{attribute 'qualified_only'}
VAR_GLOBAL CONSTANT
	//This GVL contains a list of TwinCAT Errors and their corresponding error codes.
	MAX_INDEX		: INT := 744;
	
	{warning disable C0198} //disable string length warning, strings will automatically be truncated
	List			: ARRAY[0..MAX_INDEX] OF ST_TcError :=
	[
		//0 -----------------------------------
		(code		:= 0
		,message 	:= '0.  No Error')
		//1 -----------------------------------
		,(code		:= 1
		,message 	:= '1.  Internal error')
		//2 -----------------------------------
		,(code		:= 2
		,message 	:= '2.  No Rtime')
		//3 -----------------------------------
		,(code		:= 3
		,message 	:= '3.  Allocation locked memory error')
		//4 -----------------------------------
		,(code		:= 4
		,message 	:= '4.  Insert mailbox error')
		//5 -----------------------------------
		,(code		:= 5
		,message 	:= '5.  Wrong receive HMSG')
		//6 -----------------------------------
		,(code		:= 6
		,message 	:= '6.  target port not found')
		//7 -----------------------------------
		,(code		:= 7
		,message 	:= '7.  target machine not found')
		//8 -----------------------------------
		,(code		:= 8
		,message 	:= '8.  Unknown command ID')
		//9 -----------------------------------
		,(code		:= 9
		,message 	:= '9.  Bad task ID')
		//10 -----------------------------------
		,(code		:= 10
		,message 	:= '10.  No IO')
		//11 -----------------------------------
		,(code		:= 11
		,message 	:= '11.  Unknown ADS command')
		//12 -----------------------------------
		,(code		:= 12
		,message 	:= '12.  Win 32 error')
		//13 -----------------------------------
		,(code		:= 13
		,message 	:= '13.  Port not connected')
		//14 -----------------------------------
		,(code		:= 14
		,message 	:= '14.  Invalid ADS length')
		//15 -----------------------------------
		,(code		:= 15
		,message 	:= '15.  Invalid ADS Net ID')
		//16 -----------------------------------
		,(code		:= 16
		,message 	:= '16.  Low Installation level')
		//17 -----------------------------------
		,(code		:= 17
		,message 	:= '17.  No debug available')
		//18 -----------------------------------
		,(code		:= 18
		,message 	:= '18.  Port disabled')
		//19 -----------------------------------
		,(code		:= 19
		,message 	:= '19.  Port already connected')
		//20 -----------------------------------
		,(code		:= 20
		,message 	:= '20.  ADS Sync Win32 error')
		//21 -----------------------------------
		,(code		:= 21
		,message 	:= '21.  ADS Sync Timeout')
		//22 -----------------------------------
		,(code		:= 22
		,message 	:= '22.  ADS Sync AMS error')
		//23 -----------------------------------
		,(code		:= 23
		,message 	:= '23.  ADS Sync no index map')
		//24 -----------------------------------
		,(code		:= 24
		,message 	:= '24.  Invalid ADS port')
		//25 -----------------------------------
		,(code		:= 25
		,message 	:= '25.  No memory')
		//26 -----------------------------------
		,(code		:= 26
		,message 	:= '26.  TCP send error')
		//27 -----------------------------------
		,(code		:= 27
		,message 	:= '27.  Host unreachable')
		//28 -----------------------------------
		,(code		:= 28
		,message 	:= '28.  Invalid AMS fragment')
		//29 -----------------------------------
		,(code		:= 1280
		,message 	:= '1280.  No locked memory can be allocated')
		//30 -----------------------------------
		,(code		:= 1281
		,message 	:= '1281.  The size of the router memory could not be changed')
		//31 -----------------------------------
		,(code		:= 1282
		,message 	:= '1282.  The mailbox has reached the maximum number of possible messages. The current sent message was rejected')
		//32 -----------------------------------
		,(code		:= 1283
		,message 	:= '1283.  The mailbox has reached the maximum number of possible messages.')
		//33 -----------------------------------
		,(code		:= 1284
		,message 	:= '1284.  Unknown port type')
		//34 -----------------------------------
		,(code		:= 1285
		,message 	:= '1285.  Router is not initialized')
		//35 -----------------------------------
		,(code		:= 1286
		,message 	:= '1286.  The desired port number is already assigned')
		//36 -----------------------------------
		,(code		:= 1287
		,message 	:= '1287.  Port not registered')
		//37 -----------------------------------
		,(code		:= 1288
		,message 	:= '1288.  The maximum number of Ports reached')
		//38 -----------------------------------
		,(code		:= 1289
		,message 	:= '1289.  Invalid port')
		//39 -----------------------------------
		,(code		:= 1290
		,message 	:= '1290.  TwinCAT Router not active')
		//40 -----------------------------------
		,(code		:= 1792
		,message 	:= '1792.  error class <device error>')
		//41 -----------------------------------
		,(code		:= 1793
		,message 	:= '1793.  Service is not supported by server')
		//42 -----------------------------------
		,(code		:= 1794
		,message 	:= '1794.  invalid index group')
		//43 -----------------------------------
		,(code		:= 1795
		,message 	:= '1795.  invalid index offset')
		//44 -----------------------------------
		,(code		:= 1796
		,message 	:= '1796.  reading/writing not permitted')
		//45 -----------------------------------
		,(code		:= 1797
		,message 	:= '1797.  parameter size not correct')
		//46 -----------------------------------
		,(code		:= 1798
		,message 	:= '1798.  invalid parameter value(s)')
		//47 -----------------------------------
		,(code		:= 1799
		,message 	:= '1799.  device is not in a ready state')
		//48 -----------------------------------
		,(code		:= 1800
		,message 	:= '1800.  device is busy')
		//49 -----------------------------------
		,(code		:= 1801
		,message 	:= '1801.  invalid context (must be in Windows)')
		//50 -----------------------------------
		,(code		:= 1802
		,message 	:= '1802.  out of memory')
		//51 -----------------------------------
		,(code		:= 1803
		,message 	:= '1803.  invalid parameter value(s)')
		//52 -----------------------------------
		,(code		:= 1804
		,message 	:= '1804.  not found (files, ...)')
		//53 -----------------------------------
		,(code		:= 1805
		,message 	:= '1805.  syntax error in command or file')
		//54 -----------------------------------
		,(code		:= 1806
		,message 	:= '1806.  objects do not match')
		//55 -----------------------------------
		,(code		:= 1807
		,message 	:= '1807.  object already exists')
		//56 -----------------------------------
		,(code		:= 1808
		,message 	:= '1808.  symbol not found')
		//57 -----------------------------------
		,(code		:= 1809
		,message 	:= '1809.  symbol version invalid')
		//58 -----------------------------------
		,(code		:= 1810
		,message 	:= '1810.  server is in invalid state')
		//59 -----------------------------------
		,(code		:= 1811
		,message 	:= '1811.  AdsTransMode not supported')
		//60 -----------------------------------
		,(code		:= 1812
		,message 	:= '1812.  Notification handle is invalid')
		//61 -----------------------------------
		,(code		:= 1813
		,message 	:= '1813.  Notification client not registered')
		//62 -----------------------------------
		,(code		:= 1814
		,message 	:= '1814.  no more notification handles')
		//63 -----------------------------------
		,(code		:= 1815
		,message 	:= '1815.  size for watch too big')
		//64 -----------------------------------
		,(code		:= 1816
		,message 	:= '1816.  device not initialized')
		//65 -----------------------------------
		,(code		:= 1817
		,message 	:= '1817.  device has a timeout')
		//66 -----------------------------------
		,(code		:= 1818
		,message 	:= '1818.  query interface failed')
		//67 -----------------------------------
		,(code		:= 1819
		,message 	:= '1819.  wrong interface required')
		//68 -----------------------------------
		,(code		:= 1820
		,message 	:= '1820.  class ID is invalid')
		//69 -----------------------------------
		,(code		:= 1821
		,message 	:= '1821.  object ID is invalid')
		//70 -----------------------------------
		,(code		:= 1822
		,message 	:= '1822.  request is pending')
		//71 -----------------------------------
		,(code		:= 1823
		,message 	:= '1823.  request is aborted')
		//72 -----------------------------------
		,(code		:= 1824
		,message 	:= '1824.  signal warning')
		//73 -----------------------------------
		,(code		:= 1825
		,message 	:= '1825.  invalid array index')
		//74 -----------------------------------
		,(code		:= 1826
		,message 	:= '1826.  symbol not active')
		//75 -----------------------------------
		,(code		:= 1827
		,message 	:= '1827.  access denied')
		//76 -----------------------------------
		,(code		:= 1828
		,message 	:= '1828.  missing license')
		//77 -----------------------------------
		,(code		:= 1829
		,message 	:= '1829.  license expired')
		//78 -----------------------------------
		,(code		:= 1830
		,message 	:= '1830.  license exceeded')
		//79 -----------------------------------
		,(code		:= 1831
		,message 	:= '1831.  license invalid')
		//80 -----------------------------------
		,(code		:= 1832
		,message 	:= '1832.  license invalid system id')
		//81 -----------------------------------
		,(code		:= 1833
		,message 	:= '1833.  license not time limited')
		//82 -----------------------------------
		,(code		:= 1834
		,message 	:= '1834.  license issue time in the future')
		//83 -----------------------------------
		,(code		:= 1835
		,message 	:= '1835.  license time period to long')
		//84 -----------------------------------
		,(code		:= 1836
		,message 	:= '1836.  exception occured during system start')
		//85 -----------------------------------
		,(code		:= 1837
		,message 	:= '1837.  License file read twice')
		//86 -----------------------------------
		,(code		:= 1838
		,message 	:= '1838.  invalid signature')
		//87 -----------------------------------
		,(code		:= 1839
		,message 	:= '1839.  public key certificate')
		//88 -----------------------------------
		,(code		:= 1856
		,message 	:= '1856.  Error class <client error>')
		//89 -----------------------------------
		,(code		:= 1857
		,message 	:= '1857.  invalid parameter at service')
		//90 -----------------------------------
		,(code		:= 1858
		,message 	:= '1858.  polling list is empty')
		//91 -----------------------------------
		,(code		:= 1859
		,message 	:= '1859.  var connection already in use')
		//92 -----------------------------------
		,(code		:= 1860
		,message 	:= '1860.  invoke ID in use')
		//93 -----------------------------------
		,(code		:= 1861
		,message 	:= '1861.  timeout elapsed')
		//94 -----------------------------------
		,(code		:= 1862
		,message 	:= '1862.  error in win32 subsystem')
		//95 -----------------------------------
		,(code		:= 1863
		,message 	:= '1863.  Invalid client timeout value')
		//96 -----------------------------------
		,(code		:= 1864
		,message 	:= '1864.  ads-port not opened')
		//97 -----------------------------------
		,(code		:= 1872
		,message 	:= '1872.  internal error in ads sync')
		//98 -----------------------------------
		,(code		:= 1873
		,message 	:= '1873.  hash table overflow')
		//99 -----------------------------------
		,(code		:= 1874
		,message 	:= '1874.  key not found in hash')
		//100 -----------------------------------
		,(code		:= 1875
		,message 	:= '1875.  no more symbols in cache')
		//101 -----------------------------------
		,(code		:= 1876
		,message 	:= '1876.  invalid response received')
		//102 -----------------------------------
		,(code		:= 1877
		,message 	:= '1877.  sync port is locked')
		//103 -----------------------------------
		,(code		:= 4096
		,message 	:= '4096.  Internal fatal error in the TwinCAT real-time system')
		//104 -----------------------------------
		,(code		:= 4097
		,message 	:= '4097.  Timer value not vaild')
		//105 -----------------------------------
		,(code		:= 4098
		,message 	:= '4098.  Task pointer has the invalid value ZERO')
		//106 -----------------------------------
		,(code		:= 4099
		,message 	:= '4099.  Task stack pointer has the invalid value ZERO')
		//107 -----------------------------------
		,(code		:= 4100
		,message 	:= '4100.  The demand task priority is already assigned')
		//108 -----------------------------------
		,(code		:= 4101
		,message 	:= '4101.  No more free TCB (Task Control Block) available. Maximum number of TCBs is 64')
		//109 -----------------------------------
		,(code		:= 4102
		,message 	:= '4102.  No more free semaphores available. Maximum number of semaphores is 64')
		//110 -----------------------------------
		,(code		:= 4103
		,message 	:= '4103.  No more free queue available. Maximum number of queue is 64')
		//111 -----------------------------------
		,(code		:= 4109
		,message 	:= '4109.  An external synchronization interrupt is already applied')
		//112 -----------------------------------
		,(code		:= 4110
		,message 	:= '4110.  No external synchronization interrupt applied')
		//113 -----------------------------------
		,(code		:= 4111
		,message 	:= '4111.  The apply of the external synchronization interrupt failed')
		//114 -----------------------------------
		,(code		:= 4112
		,message 	:= '4112.  Call of a service function in the wrong context')
		//115 -----------------------------------
		,(code		:= 4119
		,message 	:= '4119.  Intel VT-x extension is not supported')
		//116 -----------------------------------
		,(code		:= 4120
		,message 	:= '4120.  Intel VT-x extension is not enabled in system BIOS')
		//117 -----------------------------------
		,(code		:= 4121
		,message 	:= '4121.  Missing function in Intel VT-x extension')
		//118 -----------------------------------
		,(code		:= 4122
		,message 	:= '4122.  Enabling Intel VT-x fails')
		//119 -----------------------------------
		,(code		:= 10060
		,message 	:= '10060.  A connection attempt failed because the connected party did not properly respond after a period of time, or established connection failed because connected host has failed to respond.')
		//120 -----------------------------------
		,(code		:= 10061
		,message 	:= '10061.  No connection could be made because the target machine actively refused it. This error normally occurs when you try to connect to a service which is inactive on a different host - a service without a server application.')
		//121 -----------------------------------
		,(code		:= 10065
		,message 	:= '10065.  No route to a host. A socket operation was attempted to an unreachable host')
		//122 -----------------------------------
		,(code		:= 16384
		,message 	:= '16384.  Internal error Internal system error in the NC on ring 0, no further details.')
		//123 -----------------------------------
		,(code		:= 16385
		,message 	:= '16385.  Memory error The ring-0 memory management is not providing the required memory. This is usually a result of another error, as a result of which the controller will halt normal operation (now if not before).')
		//124 -----------------------------------
		,(code		:= 16386
		,message 	:= '16386.  Nc retain data error (persistent data) Error while loading the Nc retain data. The axes concerned are no longer referenced (status flag Homed is set to FALSE).')
		//125 -----------------------------------
		,(code		:= 16400
		,message 	:= '16400.  Channel identifier not allowed Either an unacceptable value (not 1...255) has been used, or a channel that does not exist in the system has been named.')
		//126 -----------------------------------
		,(code		:= 16401
		,message 	:= '16401.  Group identifier not allowed Either an unacceptable value (not 1...255) has been used, or a group that does not exist in the system has been named.')
		//127 -----------------------------------
		,(code		:= 16402
		,message 	:= '16402.  Axis identifier not allowed Either an unacceptable value (not 1...255) has been used, or an axis that does not exist in the system has been named.')
		//128 -----------------------------------
		,(code		:= 16403
		,message 	:= '16403.  Encoder identifier not allowed Either an unacceptable value (not 1...255) has been used, or a encoder that does not exist in the system has been named.')
		//129 -----------------------------------
		,(code		:= 16404
		,message 	:= '16404.  Controller identifier not allowed Either an unacceptable value (not 1...255) has been used, or a controller that does not exist in the system has been named.')
		//130 -----------------------------------
		,(code		:= 16405
		,message 	:= '16405.  Drive identifier not allowed Either an unacceptable value (not 1...255) has been used, or a drive that does not exist in the system has been named.')
		//131 -----------------------------------
		,(code		:= 16406
		,message 	:= '16406.  Table identifier not allowed Either an unacceptable value (not 1...255) has been used, or a table that does not exist in the system has been named.')
		//132 -----------------------------------
		,(code		:= 16416
		,message 	:= '16416.  No process image No PLC-axis interface during creation of an axis.')
		//133 -----------------------------------
		,(code		:= 16417
		,message 	:= '16417.  No process image No axis-PLC interface during creation of an axis.')
		//134 -----------------------------------
		,(code		:= 16418
		,message 	:= '16418.  No process image No encoder-I/O interface during creation of an axis.')
		//135 -----------------------------------
		,(code		:= 16419
		,message 	:= '16419.  No process image No I/O-encoder interface during creation of an axis.')
		//136 -----------------------------------
		,(code		:= 16420
		,message 	:= '16420.  No process image No drive-I/O interface during creation of an axis.')
		//137 -----------------------------------
		,(code		:= 16421
		,message 	:= '16421.  No process image No I/O-drive interface during creation of an axis.')
		//138 -----------------------------------
		,(code		:= 16432
		,message 	:= '16432.  Coupling type not allowed Unacceptable master/slave coupling type.')
		//139 -----------------------------------
		,(code		:= 16433
		,message 	:= '16433.  Axis type not allowed Unacceptable type specification during creation of an axis.')
		//140 -----------------------------------
		,(code		:= 16448
		,message 	:= '16448.  Axis is incompatible Axis is not suitable for the intended purpose. A high speed/low speed axis, for example, cannot function as a slave in an axis coupling.')
		//141 -----------------------------------
		,(code		:= 16464
		,message 	:= '16464.  Channel not ready for operation The channel is not complete, and is therefore not ready for operation. This is usually a consequence of problems at system start-up.')
		//142 -----------------------------------
		,(code		:= 16465
		,message 	:= '16465.  Group not ready for operation The group is not complete, and is therefore not ready for operation. This is usually a consequence of problems at system start-up.')
		//143 -----------------------------------
		,(code		:= 16466
		,message 	:= '16466.  Axis not ready for operation The axis is not complete, and is therefore not ready for operation. This is usually a consequence of problems at system start-up.')
		//144 -----------------------------------
		,(code		:= 16480
		,message 	:= '16480.  Channel exists The channel that is to be created already exists.')
		//145 -----------------------------------
		,(code		:= 16481
		,message 	:= '16481.  Group exists The group that is to be created already exists.')
		//146 -----------------------------------
		,(code		:= 16482
		,message 	:= '16482.  Axis exists The axis that is to be created already exists.')
		//147 -----------------------------------
		,(code		:= 16483
		,message 	:= '16483.  Table exists The table that is to be created already exists, resp. it is tried internally to use an already existing table id ( e.g. for the universal flying saw).')
		//148 -----------------------------------
		,(code		:= 16496
		,message 	:= '16496.  Axis index not allowed The location within the channel specified for an axis is not allowed.')
		//149 -----------------------------------
		,(code		:= 16497
		,message 	:= '16497.  Axis index not allowed The location within the group specified for an axis is not allowed.')
		//150 -----------------------------------
		,(code		:= 16641
		,message 	:= '16641.  Group index not allowed The location within the channel specified for an group is not allowed.')
		//151 -----------------------------------
		,(code		:= 16642
		,message 	:= '16642.  Null pointer The pointer to the group is invalid. This is usually a consequence of an error at system start-up.')
		//152 -----------------------------------
		,(code		:= 16643
		,message 	:= '16643.  No process image It is not possible to exchange data with the PLC. Possible causes: n The channel does not have an interface (no interpreter present) n The connection to the PLC is faulty')
		//153 -----------------------------------
		,(code		:= 16644
		,message 	:= '16644.  M-function index not allowed Unacceptable M-function (not 0...159) detected at the execution level.')
		//154 -----------------------------------
		,(code		:= 16645
		,message 	:= '16645.  No memory No more system memory is available. This is usually the result of another error.')
		//155 -----------------------------------
		,(code		:= 16646
		,message 	:= '16646.  Not ready The function is not presently available, because a similar function is already being processed. This is usually the result of access conflicts: more than one instance wants to issue commands to the channel. This can, for example, be the consequence of an incorrect PLC program.')
		//156 -----------------------------------
		,(code		:= 16647
		,message 	:= '16647.  Function/command not supported A requested function or command is not supported by the channel.')
		//157 -----------------------------------
		,(code		:= 16648
		,message 	:= '16648.  Invalid parameter while starting Parameters to start the channel (TwinCAT-Start) are invalid. Typically there is an invalid memory size or channel type requested.')
		//158 -----------------------------------
		,(code		:= 16649
		,message 	:= '16649.  Channel function/command not executable A channel function e.g. interpreter start is not executable because the channel is already busy, no program is loaded or in an error state.')
		//159 -----------------------------------
		,(code		:= 16650
		,message 	:= '16650.  ItpGoAhead not executable The requested command is not executable, because the interpreter is not executing a dekoder stop.')
		//160 -----------------------------------
		,(code		:= 16656
		,message 	:= '16656.  Error opening a file The specified file does not exist. Example: NC program unknown.')
		//161 -----------------------------------
		,(code		:= 16657
		,message 	:= '16657.  Syntax error during loading The NC has found a syntax error when loading an NC program.')
		//162 -----------------------------------
		,(code		:= 16658
		,message 	:= '16658.  Syntax error during interpretation The NC has found a syntax error when executing an NC program.')
		//163 -----------------------------------
		,(code		:= 16659
		,message 	:= '16659.  Missing subroutine The NC has found a missing subroutine while loading.')
		//164 -----------------------------------
		,(code		:= 16660
		,message 	:= '16660.  Loading buffer of interpreter is too small The capacity of the interpreter loading buffer has been exceeded.')
		//165 -----------------------------------
		,(code		:= 16661
		,message 	:= '16661.  ?Symbolic?  - reserved')
		//166 -----------------------------------
		,(code		:= 16662
		,message 	:= '16662.  ?Symbolic?  - reserved')
		//167 -----------------------------------
		,(code		:= 16663
		,message 	:= '16663.  ?Subroutine incomplete?  Header of subroutine is missing')
		//168 -----------------------------------
		,(code		:= 16672
		,message 	:= '16672.  Divide by zero The NC encountered a computation error during execution: division by 0.')
		//169 -----------------------------------
		,(code		:= 16673
		,message 	:= '16673.  Invalid circle parameterisation The NC encountered a computation error during execution: The specified circle cannot be calculated.')
		//170 -----------------------------------
		,(code		:= 16674
		,message 	:= '16674.  ?Invalid FPU-Operation? The NC encountered an invalid FPU-Operation during exectuion. This error occurs e.g. by calculating the square root of a negative number.')
		//171 -----------------------------------
		,(code		:= 16688
		,message 	:= '16688.  Stack overflow: subroutines The NC encountered a stack overflow during execution: too many subroutine levels.')
		//172 -----------------------------------
		,(code		:= 16689
		,message 	:= '16689.  Stack underflow: subroutines The NC encountered a stack underflow during execution: too many subroutine return commands. Note: A main program must not end with a return command.')
		//173 -----------------------------------
		,(code		:= 16690
		,message 	:= '16690.  Stack overflow: arithmetic unit The NC encountered a stack overflow during execution: The calculation is too complex, or has not been correctly written.')
		//174 -----------------------------------
		,(code		:= 16691
		,message 	:= '16691.  Stack underflow: arithmetic unit The NC encountered a stack underflow during execution: The calculation is too complex, or has not been correctly written.')
		//175 -----------------------------------
		,(code		:= 16704
		,message 	:= '16704.  Register index not allowed The NC encountered an unacceptable register index during execution: Either the program contains an unacceptable value (not R0...R999) or a pointer register contains an unacceptable value.')
		//176 -----------------------------------
		,(code		:= 16705
		,message 	:= '16705.  Unacceptable G-function index The NC has encountered an unacceptable G-function (not 0...159) during execution.')
		//177 -----------------------------------
		,(code		:= 16706
		,message 	:= '16706.  Unacceptable M-function index The NC has encountered an unacceptable M-function (not 0...159) during execution.')
		//178 -----------------------------------
		,(code		:= 16707
		,message 	:= '16707.  Unacceptable extended address The NC has encountered an unacceptable extended address (not 1...9) during execution.')
		//179 -----------------------------------
		,(code		:= 16708
		,message 	:= '16708.  Unacceptable index to the internal H-function The NC has encountered an unacceptable internal H-function in the course of processing. This is usually a consequence of an error during loading.')
		//180 -----------------------------------
		,(code		:= 16709
		,message 	:= '16709.  Machine data value unacceptable While processing instructions the NC has detected an impermissible value for the machine data (MDB) (not 0?7).')
		//181 -----------------------------------
		,(code		:= 16720
		,message 	:= '16720.  Cannot change tool params here The NC has encountered an unacceptable change of parameters for the tool compensation during execution. This error occured for instance by changing the tool radius and programming a circle in the same block.')
		//182 -----------------------------------
		,(code		:= 16721
		,message 	:= '16721.  Cannot calculate tool compensation The NC has encountered an error by  the calculation of the tool compensation')
		//183 -----------------------------------
		,(code		:= 16722
		,message 	:= '16722.  Tool compensation: The plane for the tool compensation cannot be changed here. This error occured for instance by changing the tool plane when the compensation is turned on or active.')
		//184 -----------------------------------
		,(code		:= 16723
		,message 	:= '16723.  Tool compensation:  The D-Word is missing or invalid by turning on the tool compensation.')
		//185 -----------------------------------
		,(code		:= 16724
		,message 	:= '16724.  Tool compensation:  The spezified tool radius is invalid because the value is less or equal zero.')
		//186 -----------------------------------
		,(code		:= 16725
		,message 	:= '16725.  Tool compensation: The tool radius cannot be changed here')
		//187 -----------------------------------
		,(code		:= 16726
		,message 	:= '16726.  Tool compensation:  Collision Detection Table is full.')
		//188 -----------------------------------
		,(code		:= 16727
		,message 	:= '16727.  Tool compensation: Internal error while turning on the contour collision detection.')
		//189 -----------------------------------
		,(code		:= 16728
		,message 	:= '16728.  Tool compensation:  Internal error within the contour collision detection - update reversed geo failed.')
		//190 -----------------------------------
		,(code		:= 16729
		,message 	:= '16729.  Tool compensation:  Unexpected combination of geometrie types by active contour collision detection.')
		//191 -----------------------------------
		,(code		:= 16730
		,message 	:= '16730.  Tool compensation: Programmed inner circle is smaller than the cutter radius')
		//192 -----------------------------------
		,(code		:= 16731
		,message 	:= '16731.  Tool compensation:  Bottle neck detection recognized contour violation')
		//193 -----------------------------------
		,(code		:= 16732
		,message 	:= '16732.  Table for corrected entries is full')
		//194 -----------------------------------
		,(code		:= 16733
		,message 	:= '16733.  Input table for tangential following is full')
		//195 -----------------------------------
		,(code		:= 16734
		,message 	:= '16734.  Executing table for tangential following is full')
		//196 -----------------------------------
		,(code		:= 16735
		,message 	:= '16735.  Geometric entry for tangential following can not be calculated')
		//197 -----------------------------------
		,(code		:= 16736
		,message 	:= '16736.  reserved')
		//198 -----------------------------------
		,(code		:= 16737
		,message 	:= '16737.  reserved')
		//199 -----------------------------------
		,(code		:= 16738
		,message 	:= '16738.  The acutal active interpolation rules (g-code), zero-shifts, or rotation cannot be detected')
		//200 -----------------------------------
		,(code		:= 16752
		,message 	:= '16752.  Error while loading: Invalid parameter The NC has found an invalid parameter while loading an NC program.')
		//201 -----------------------------------
		,(code		:= 16753
		,message 	:= '16753.  Invalid contour start position The NC encountered a computation error during execution: The specified contour cannot be calculated because the initial position is not on the contour.')
		//202 -----------------------------------
		,(code		:= 16754
		,message 	:= '16754.  Retrace: Invalid internal entry index The NC encountered an invalid internal entry index during execution of the retrace function.')
		//203 -----------------------------------
		,(code		:= 16896
		,message 	:= '16896.  Group ID not allowed The value for the group ID is not allowed, e.g. because it has already been assigned, is less than or equal to zero, or is greater than 255.')
		//204 -----------------------------------
		,(code		:= 16897
		,message 	:= '16897.  Group type not allowed The value for the group type is unacceptable because it is not defined. Type 1: PTP group with slaves (servo) Type 5: DXD group with slaves (3D group) Type 6: High/low speed group Type 7: Stepper motor group Type 8: 0D group')
		//205 -----------------------------------
		,(code		:= 16898
		,message 	:= '16898.  Master axis index not allowed  The value for the master axis index in an interpolating 3D group is not allowed, because, for instance, it has gone outside the value range. Index 0: X axis (first master axis) Index 1: Y axis (second master axis) Index 2: Z axis (third master axis)')
		//206 -----------------------------------
		,(code		:= 16899
		,message 	:= '16899.  Slave axis index not allowed (INTERNAL ERROR) The value for the slave axis index in a group is not allowed, because, for instance, it has passed outside the value range, the slave location to be used when inserting a new slave connection is already occupied, or because no slave is present when such a connection is being removed. Index 0: First slave axis Index 1: Second slave axis Index 2: etc.')
		//207 -----------------------------------
		,(code		:= 16900
		,message 	:= '16900.  (INTERNAL ERROR) GROUPERR_INTERNAL')
		//208 -----------------------------------
		,(code		:= 16901
		,message 	:= '16901.  Invalid cycle time for statement execution task (SAF) The value of the cycle time for the NC block execution task (SAF 1/2) is not allowed, because it has passed outside the value range.')
		//209 -----------------------------------
		,(code		:= 16902
		,message 	:= '16902.  GROUPERR_RANGE_MAXELEMENTSINAXIS')
		//210 -----------------------------------
		,(code		:= 16903
		,message 	:= '16903.  Invalid cycle time for the statement preparation task (SVB) The value of the cycle time for the NC statement preparation task (SVB 1/2) is not allowed, because it has passed outside the value range.')
		//211 -----------------------------------
		,(code		:= 16904
		,message 	:= '16904.  Single step mode not allowed The flag for the activation or deactivation of single step mode is not allowed. Value 0: Passive (buffered operation) Value 1: Active (single-block operation)')
		//212 -----------------------------------
		,(code		:= 16905
		,message 	:= '16905.  Group deactivation not allowed (INTERNAL ERROR) The flag for the deactivation or activation of the complete group is not allowed. Value 0: Group active Value 1: Group passive')
		//213 -----------------------------------
		,(code		:= 16906
		,message 	:= '16906.  Statement execution state (SAF state) not allowed (INTERNAL ERROR) The value for the state of the block execution state machine (SAF state) is not allowed. This error occurs on passing outside the range of values, or if the state machine enters an error state.')
		//214 -----------------------------------
		,(code		:= 16907
		,message 	:= '16907.  Channel address The group does not have a channel, or the channel address has not been initialised.')
		//215 -----------------------------------
		,(code		:= 16908
		,message 	:= '16908.  Axis address (master axis) The group does not have a master axis (or axes) or the axis address(es) has (have) not been initialised.')
		//216 -----------------------------------
		,(code		:= 16909
		,message 	:= '16909.  Master axis address A new master/slave coupling is to be inserted into the group, but there is no valid address for the leading master axis.')
		//217 -----------------------------------
		,(code		:= 16910
		,message 	:= '16910.  Slave axis address A master/slave coupling is to be inserted into the group, but there is no valid address for the slave axis.')
		//218 -----------------------------------
		,(code		:= 16911
		,message 	:= '16911.  Slave set value generator address A master/slave coupling is to be inserted into the group, but there is no valid address for the slave set value generator.')
		//219 -----------------------------------
		,(code		:= 16912
		,message 	:= '16912.  Encoder address An axis in the group does not have an encoder, or the encoder address has not been initialised.')
		//220 -----------------------------------
		,(code		:= 16913
		,message 	:= '16913.  Controller address An axis in the group does not have a controller, or the controller address has not been initialised.')
		//221 -----------------------------------
		,(code		:= 16914
		,message 	:= '16914.  Drive address An axis in the group does not have a drive, or the drive address has not been initialised.')
		//222 -----------------------------------
		,(code		:= 16915
		,message 	:= '16915.  GROUPERR_ADDR_MASTERGENERATOR')
		//223 -----------------------------------
		,(code		:= 16916
		,message 	:= '16916.  Axis interface NC to PLC address Group/axis does not have an axis interface from the NC to the PLC, or the axis interface address has not been initialised.')
		//224 -----------------------------------
		,(code		:= 16917
		,message 	:= '16917.  Slave axis address An existing master/slave coupling is to be removed from the group, but there is no valid address for the slave axis.')
		//225 -----------------------------------
		,(code		:= 16918
		,message 	:= '16918.  ?Table adress unknown? The table, respectively the table ID, is unknown. This table is used for the master/slave coupling or for the characteristic curve.')
		//226 -----------------------------------
		,(code		:= 16919
		,message 	:= '16919.  NcControl address The NcControl address has not been initialised.')
		//227 -----------------------------------
		,(code		:= 16920
		,message 	:= '16920.  Axis is blocked for commands while persistent NC data are queued Axis is blocked for commands while waiting for valid IO data to accept the queued persistent NC data.')
		//228 -----------------------------------
		,(code		:= 16921
		,message 	:= '16921.  The scaling mode MASTER-AUTOOFFSET is invalid because no reference table was found. The used scaling mode MASTER-AUTOOFFSET is invalid in this context because an existing reference table is missing.')
		//229 -----------------------------------
		,(code		:= 16922
		,message 	:= '16922.  The master axis start position does not permit synchronisation When a slave axis is being coupled on, the position of the master axis does not permit synchronisation at the given synchronisation positions.')
		//230 -----------------------------------
		,(code		:= 16923
		,message 	:= '16923.  Slave coupling factor (gearing factor) of 0.0 is not allowed A master/slave coupling with a gearing factor of 0.0 is being created. This value is not allowed, since it does not correspond to any possible coupling, and division will generate an FPU exception.')
		//231 -----------------------------------
		,(code		:= 16924
		,message 	:= '16924.  Insertion of master axis into group not allowed  A master axis is to be inserted into a group at a location that is already occupied by another master axis.')
		//232 -----------------------------------
		,(code		:= 16925
		,message 	:= '16925.  Deletion of master axis from group not allowed (INTERNAL ERROR) A master axis is to be removed from a location in a group that is not in fact occupied by master axis.')
		//233 -----------------------------------
		,(code		:= 16926
		,message 	:= '16926.  ?Function/feature is not supported from the setpoint generator A function or feature is not supported from the setpoint generator (e.g. PTP master setpoint generator). This can be in general or only in a special situation.')
		//234 -----------------------------------
		,(code		:= 16927
		,message 	:= '16927.  Group initialisation Group has not been initialised. Although the group has been created, the rest of the initialisation has not been performed (1. Initialisation of group I/O, 2. Initialisation of group, 3. Reset group).')
		//235 -----------------------------------
		,(code		:= 16928
		,message 	:= '16928.  Group not ready / group not ready for new task The group is being given a new task while it is still in the process of executing an existing task. This request is not allowed because it would interrupt the execution of the previous task. The new task could, for instance, be a positioning command, or the set actual position function. Precisely the converse relationships apply for the set new end position function. In that case, the group/axis must still be actively moving in order to be able to cause a change in the end position.')
		//236 -----------------------------------
		,(code		:= 16929
		,message 	:= '16929.  Requested set velocity is not allowed The value requested for the set velocity of a positioning task is less than or equal to zero, larger than the maximum velocity (see axis parameters), or, in the case of servo-drives, is larger than the reference velocity of the axis (see drive parameters).')
		//237 -----------------------------------
		,(code		:= 16930
		,message 	:= '16930.  Requested target position is not allowed (master axis) The requested value for the target position of a positioning task is not within the software end locations. In other words, it is either less than the minimum software end location or larger than the maximum software end location. This check is only carried out if the relevant end position monitoring is active.')
		//238 -----------------------------------
		,(code		:= 16931
		,message 	:= '16931.  No enable for controller and/or feed (Master axis) The axis enables for the master axis needed for positioning are not present. This can involve the controller enable and/or the relevant, direction-dependent feed enable (see axis interface PLC®NC).')
		//239 -----------------------------------
		,(code		:= 16932
		,message 	:= '16932.  Movement smaller than one encoder increment (INTERNAL ERROR) The distance that a group/axis is supposed to move is smaller than the physical significance of one encoder increment. In other words the movement is smaller than the scaling factor of the axis. The reaction to this is that the axis is reported as having logically finished without having actively moved. This means that an external error is not generated for the user. This error is also issued for high/low speed axes if a loop movement with non-zero parameters is smaller than the sum of the creeping and braking distances. In such a case it is not meaningful to either exceed or to fail to reach the target position.')
		//240 -----------------------------------
		,(code		:= 16933
		,message 	:= '16933.  Drive not ready during axis start During an axis start it is ascertained that the drive is not ready. The following are possible causes: - the drive is in failure state (hardware fault) - the drive is in the starting-up stage (e.g. following an axis reset preceded by a hardware fault) - the drive has not been enabled Remark: The time required for booting a drive after a hardware fault can amount to several seconds.')
		//241 -----------------------------------
		,(code		:= 16934
		,message 	:= '16934.  Invalid parameters of the emergency stop. The parameter of the E-Stop are invalid. Either the deceleration and the jerk are less than zero or one of the parameters is weaker than the corresponding parameter of the start data.')
		//242 -----------------------------------
		,(code		:= 16935
		,message 	:= '16935.  The setpoint generator is inactive such that no instructions are accepted.')
		//243 -----------------------------------
		,(code		:= 16936
		,message 	:= '16936.  ?Requested traverse distance is not allowed? The requested traverse distance or looping distance is smaller than the braking distance of the two/speed axis.')
		//244 -----------------------------------
		,(code		:= 16937
		,message 	:= '16937.  Requested target position is not allowed (slave axis) The value for the target position of a positioning task when calculated for the slave axis is not within the software end locations. In other words, it is either less than the minimum software end location or larger than the maximum software end location. This check is only carried out if the relevant end position monitoring is active.')
		//245 -----------------------------------
		,(code		:= 16938
		,message 	:= '16938.  No enable for controller and/or feed (slave axis) The axis enables for one or more coupled slave axes needed for positioning are not present. This can involve the controller enable and/or the relevant, direction-dependent feed enable (see axis interface PLC®NC).')
		//246 -----------------------------------
		,(code		:= 16939
		,message 	:= '16939.  The activation position (position threshold) is out of range of the actual positioning')
		//247 -----------------------------------
		,(code		:= 16940
		,message 	:= '16940.  The start or activation data of the external setpoint generation are not valid?This may be caused through:')
		//248 -----------------------------------
		,(code		:= 16941
		,message 	:= '16941.  ?Velocity is not constant? For changing the dynamic parameter acceleration und deceleration the axis has to be in dynamic state without acceleration and deceleration (that means constant velocity).')
		//249 -----------------------------------
		,(code		:= 16942
		,message 	:= '16942.  Jerk less than or equal to 0.0 is not allowed A value less than or equal to 0.0 for the jerk (PTP and CNC) is not allowed, since the jerk is by definition positive, and with a jerk of 0.0, division will generate an FPU exception.')
		//250 -----------------------------------
		,(code		:= 16943
		,message 	:= '16943.  Acceleration less than or equal to 0.0 is not allowed A value less than or equal to 0.0 for the acceleration (PTP and CNC) is not allowed, since the acceleration is positive by definition, and an acceleration of 0.0 will not allow a motion to be generated.')
		//251 -----------------------------------
		,(code		:= 16944
		,message 	:= '16944.  Absolute deceleration value less than or equal to 0.0 is not allowed A value less than or equal to 0.0 for the absolute value of the deceleration (PTP and CNC) is not allowed, since the absolute value of the deceleration is positive by definition, and an absolute value of the deceleration of 0.0 will not allow a motion to be generated.')
		//252 -----------------------------------
		,(code		:= 16945
		,message 	:= '16945.  Set velocity less than or equal to 0.0 is not allowed A value less than or equal to 0.0 or outside the range from 10-3 up to 10+10 for the set velocity (PTP and CNC) is not allowed, since the set velocity is by definition strictly positive, and with a set velocity of 0.0, division will generate an FPU exception.')
		//253 -----------------------------------
		,(code		:= 16946
		,message 	:= '16946.  ?Loss of precision when trying a positioning? The positioning is so long in space or time that decimal parts loose there relevance LOSS_OF_PRECISION).')
		//254 -----------------------------------
		,(code		:= 16947
		,message 	:= '16947.  Cycle time less than or equal to 0.0 is not allowed A value less than or equal to 0.0 for the cycle time (PTP and CNC) is not allowed, since the cycle time is by definition strictly positive, and with a cycle time of 0.0, division will generate an FPU exception.')
		//255 -----------------------------------
		,(code		:= 16948
		,message 	:= '16948.  PTP data type <intasdouble> range exceeded Such extreme parameters have been supplied for the start task, the override or the new target position that the internal data type loses its precision.')
		//256 -----------------------------------
		,(code		:= 16949
		,message 	:= '16949.  PTP LHL velocity profile cannot be generated (INTERNAL ERROR) Such extreme parameters have been supplied for the start task, the override or the new target position that it is not possible to generate a velocity profile of the type LHL (Low-High-Low).')
		//257 -----------------------------------
		,(code		:= 16950
		,message 	:= '16950.  PTP HML velocity profile cannot be generated (INTERNAL ERROR) Such extreme parameters have been supplied for the override or the new target position that it is not possible to generate a velocity profile of the type HML (High-Middle-Low).')
		//258 -----------------------------------
		,(code		:= 16951
		,message 	:= '16951.  Start data address is invalid The address of the start data is invalid.')
		//259 -----------------------------------
		,(code		:= 16952
		,message 	:= '16952.  Velocity override (start override) is not allowed The value for the velocity override is not allowed, because it is less than 0.0% or more than 100.0% (see axis interface PlcToNc). Here, 100.0 % corresponds to the integral value 1000000 in the axis interface. Value range: [0 ... 1000000]')
		//260 -----------------------------------
		,(code		:= 16953
		,message 	:= '16953.  Start type not allowed The start type supplied does not exist.')
		//261 -----------------------------------
		,(code		:= 16954
		,message 	:= '16954.  Velocity overflow (overshoot in the velocity) The new dynamic with the parameterized jerk is so weak that a velocity overflow will occur (overshoot in the velocity). The command is therefore not supported.')
		//262 -----------------------------------
		,(code		:= 16955
		,message 	:= '16955.  Start parameter for the axis structure is invalid External or internal parameters for the start structure for a positioning task are invalid. Thus, for instance, the scaling factor, the SAF cycle time or the requested velocity may be less than or equal to zero, which is not allowed.')
		//263 -----------------------------------
		,(code		:= 16956
		,message 	:= '16956.  Override generator initialisation parameter invalid One of the override generator (re)initialisation parameters is invalid.')
		//264 -----------------------------------
		,(code		:= 16957
		,message 	:= '16957.  Slave axis has not set value generator (INTERNAL ERROR) It is found that a slave axis within a group does not have a valid slave generator (set value generator). A slave axis and a slave set value generator must always be present as a pair. This is an internal error.')
		//265 -----------------------------------
		,(code		:= 16958
		,message 	:= '16958.  Table is empty Either the SVB table or the SAF table does not contain any entries.')
		//266 -----------------------------------
		,(code		:= 16959
		,message 	:= '16959.  Table is full The SVB table or the SAF table has no more free lines.')
		//267 -----------------------------------
		,(code		:= 16960
		,message 	:= '16960.  No memory available SVB memory allocation for dynamic entry in SAF table failed.')
		//268 -----------------------------------
		,(code		:= 16961
		,message 	:= '16961.  Table already contains an entry(INTERNAL ERROR) SAF table entry abandoned, because, incorrectly, an entry already exists.')
		//269 -----------------------------------
		,(code		:= 16962
		,message 	:= '16962.  Stop is already active The stop instruction is not forwarded, because it has already been activated.')
		//270 -----------------------------------
		,(code		:= 16963
		,message 	:= '16963.  Compensation has not been carried out over the full compensation sectionThe compensations start parameters do not permit compensation over the full section to be compensated. For this reason the compensation will be carried out over a smaller section.')
		//271 -----------------------------------
		,(code		:= 16964
		,message 	:= '16964.  Start parameter address for the compensation invalid (INTERNAL ERROR)Invalid address.')
		//272 -----------------------------------
		,(code		:= 16965
		,message 	:= '16965.  Compensation active Start of compensation refused, because compensation is already active.  Its also possible that the M/S axes are not active moved. Therefore an execution of the compensation is impossible.')
		//273 -----------------------------------
		,(code		:= 16966
		,message 	:= '16966.  Compensation not active Stop of compensation refused, because compensation is not active.')
		//274 -----------------------------------
		,(code		:= 16967
		,message 	:= '16967.  Compensation type invalid The type supplied for the section compensation is invalid. At the present time only compensation type 1 (trapezoidal velocity profile) is allowed.')
		//275 -----------------------------------
		,(code		:= 16968
		,message 	:= '16968.  Axis address for compensation invalid (INTERNAL ERROR) The address of the master of slave axis on which the section compensation is to act is invalid. This is an internal error.')
		//276 -----------------------------------
		,(code		:= 16969
		,message 	:= '16969.  Invalid slave address (INTERNAL ERROR) The slave address given for on-line coupling/decoupling is invalid.')
		//277 -----------------------------------
		,(code		:= 16970
		,message 	:= '16970.  Coupling velocity invalid The velocity of what is to become the master axis is 0, which means that on-line coupling is not possible.')
		//278 -----------------------------------
		,(code		:= 16971
		,message 	:= '16971.  Coupling velocities not constant The velocity of what is to become the master axis and the velocity of what is to become the slave axis are not constant, so that on-line coupling is not possible.')
		//279 -----------------------------------
		,(code		:= 16972
		,message 	:= '16972.  Cycle time less than or equal to 0.0 is not allowed A value less than or equal to 0.0 for the cycle time (Slave) is not allowed, since the cycle time is by definition strictly positive, and with a cycle time of 0.0, division will generate an FPU exception.')
		//280 -----------------------------------
		,(code		:= 16973
		,message 	:= '16973.  Decoupling task not allowed The slave axis is of such a type (e.g. a table slave) or is in such a state (master velocity 0) that on-line decoupling is not possible.')
		//281 -----------------------------------
		,(code		:= 16974
		,message 	:= '16974.  Function not allowed The function cannot logically be executed, e.g. some commands are not possible and not allowed for slave axes.')
		//282 -----------------------------------
		,(code		:= 16975
		,message 	:= '16975.  No valid table weighting has been set The weighting factor of each table is 0, so that no table can be read.')
		//283 -----------------------------------
		,(code		:= 16976
		,message 	:= '16976.  Axis type, actual position type or end position type is not allowed The start type for a positioning task in invalid. Valid start types are ABSOLUTE (1), RELATIVE (2), CONTINUOUS POSITIVE (3), CONTINUOUS NEGATIVE (4), MODULO (5), etc. . It is also possible that the types for setting a new actual position or for travel to a new end position are invalid.')
		//284 -----------------------------------
		,(code		:= 16977
		,message 	:= '16977.  Function not presently supported An NC function has been activated that is currently not released for use, or which is not even implemented. This can be a command which is not possible or not allowed for master axes.')
		//285 -----------------------------------
		,(code		:= 16978
		,message 	:= '16978.  State of state machine invalid (INTERNAL ERROR) The state of an internal state machine is invalid. This is an internal error.')
		//286 -----------------------------------
		,(code		:= 16979
		,message 	:= '16979.  Reference cam became free too soon During the referencing process for an axis it is moved in the direction of the referencing cam, and is only stopped again when the cam signal is reached. After the axis has then also physically stopped, the referencing cam must remain occupied until the axis subsequently starts back down from the cam in the normal way.')
		//287 -----------------------------------
		,(code		:= 16980
		,message 	:= '16980.  Clearance monitoring between activation of the hardware latch and appearance of the sync pulse When the clearance monitoring is active, a check is kept on whether the number of increments between activation of the hardware latch and occurrence of the sync pulse (zero pulse) has become smaller than a pre-set value. This error is generated when that happens. (See parameters for the incremental encoder)')
		//288 -----------------------------------
		,(code		:= 16981
		,message 	:= '16981.  No memory available The dynamic memory allocation for the set value generator, the SVB table or the SAF table has failed.')
		//289 -----------------------------------
		,(code		:= 16982
		,message 	:= '16982.  The table slave axis has no active table Although the table slave axis has tables, none of the tables is designated as active. If this occurs during the run time the whole master/slave group is stopped by a run time error.')
		//290 -----------------------------------
		,(code		:= 16983
		,message 	:= '16983.  Function not allowed The requested function or the requested task is not logically allowed. An example for such an error message would be set an actual position for an absolute encoder (M3000, KL5001, etc.).')
		//291 -----------------------------------
		,(code		:= 16984
		,message 	:= '16984.  Stopping compensation not allowed It is not possible to stop the compensation, since compensation is already in the stopping phase.')
		//292 -----------------------------------
		,(code		:= 16985
		,message 	:= '16985.  Slave table is being used The slave table cannot be activated, because it is currently being used.')
		//293 -----------------------------------
		,(code		:= 16986
		,message 	:= '16986.  Master or slave axis is processing a job (e.g. positioning command) while coupling is requested A master/slave coupling of a certain slave type (e.g. linear coupling) can not be executed. he master or intended slave axis is not in stand still state and is executing a job (e.g. positioning) at the same time as the coupling request received. For this couple type this is not allowed.')
		//294 -----------------------------------
		,(code		:= 16987
		,message 	:= '16987.  Slave (start) parameter is incorrect One of the slave start/coupling parameters is not allowed (Coupling factor is zero,t he master position scaling of an cam is zero, etc) .')
		//295 -----------------------------------
		,(code		:= 16988
		,message 	:= '16988.  Slave type is incorrect The slave type does not match up to the (SVB) start type.')
		//296 -----------------------------------
		,(code		:= 16989
		,message 	:= '16989.  Axis stop is already active The axis stop/Estop is not initiated, because the stop/estop is already active.')
		//297 -----------------------------------
		,(code		:= 16990
		,message 	:= '16990.  Maximum number of tables per slavegenerator reached The maximum number of tables per slave generator is reached (e.g. MC_MultiCamIn is limited to 4 tables).')
		//298 -----------------------------------
		,(code		:= 16991
		,message 	:= '16991.  The scaling mode is invalid. The used scaling is invalid in this context. Either the mode is not defined or yet not implemented or however it cannot in this constellation be put into action.')
		//299 -----------------------------------
		,(code		:= 16992
		,message 	:= '16992.  Controller enable Controller enable for the axis or for a coupled slave axis is not present (see axis interface PlcToNc). This error occurs if the controller enable is withdrawn while an axis or a group of axes (also a master/slave group) is being actively positioned. The error also occurs if a PTP axis or a coupled slave axis is started without controller enable.')
		//300 -----------------------------------
		,(code		:= 16993
		,message 	:= '16993.  Table not found No table exists with the ID prescribed or the table ID is not unique.')
		//301 -----------------------------------
		,(code		:= 16994
		,message 	:= '16994.  Incorrect table type The table referred to in the function is of the incorrect type.')
		//302 -----------------------------------
		,(code		:= 16995
		,message 	:= '16995.  Single step mode This error occurs if single step mode is selected for a group or axis and a new task is requested while one of the individual tasks is still being processed.')
		//303 -----------------------------------
		,(code		:= 16996
		,message 	:= '16996.  Group task unknown (asynchronous table entry) The group has received a task whose type or sub-type is unknown. Valid tasks can be single or multi-dimensional positioning tasks (Geo 1D, Geo 3D), referencing tasks, etc..')
		//304 -----------------------------------
		,(code		:= 16997
		,message 	:= '16997.  Group function unknown (synchronous function) The group has received a function whose type is unknown. Valid functions are Reset, Stop, New end position, Start/stop section compensation, Set actual position, Set/reset referencing status etc..')
		//305 -----------------------------------
		,(code		:= 16998
		,message 	:= '16998.  Group task for slave not allowed Group tasks are usually only possible for master axes, not for slave axes. A slave axis only moves as an indirect result of a positioning task given to its associated master axis. A slave can thus never directly be given a task.')
		//306 -----------------------------------
		,(code		:= 16999
		,message 	:= '16999.  Group function for slave not allowed Group functions are in principle only possible for master axes, not for slave axes. The only exception is represented by the Start/stop section compensation function, which is possible both for masters and for slaves. A slave cannot directly execute any other functions beyond this.')
		//307 -----------------------------------
		,(code		:= 17000
		,message 	:= '17000.  GROUPERR_GROUPFUNC_NOMOTION')
		//308 -----------------------------------
		,(code		:= 17001
		,message 	:= '17001.  ?Startposition=Setpoint Position? Invalid position parameters.')
		//309 -----------------------------------
		,(code		:= 17002
		,message 	:= '17002.  ?Parameters of the delay-denerator are invalid? Invalid external/internal parameters of the delay generator (delay time, cycle time, tics).')
		//310 -----------------------------------
		,(code		:= 17003
		,message 	:= '17003.  ?External parameters of the superimposed instruction are invalid? Invalid external parameters of the superimposed functionality (acceleration, deceleration, velocity, process velocity, length).')
		//311 -----------------------------------
		,(code		:= 17004
		,message 	:= '17004.  Invalid overridetype. The override type does not exist.')
		//312 -----------------------------------
		,(code		:= 17005
		,message 	:= '17005.  ?Activation position under/overrun? The requested activation position is located in the past of the master (e.g. when exchanging a cam table).')
		//313 -----------------------------------
		,(code		:= 17006
		,message 	:= '17006.  ?Activation impossible: Master is standing? The required activation of the correction is impossible since the master axis is  not moving.   A synchronisation is not possible, because the master axis standing and the slave axis is still not synchronous.')
		//314 -----------------------------------
		,(code		:= 17007
		,message 	:= '17007.  ?Activation mode not possible? The requested activation mode is not possible when the slave axis is moving (otherwise the slave velocity would jump to zero).')
		//315 -----------------------------------
		,(code		:= 17008
		,message 	:= '17008.  Start parameter for the compensation is invalid One of the dynamic parameters for the compensation is invalid (necessary condition): Acceleration (>0) Deceleration (>0) Process velocity (>0)')
		//316 -----------------------------------
		,(code		:= 17009
		,message 	:= '17009.  Start parameter for the compensation is invalid Velocity camber is negative.')
		//317 -----------------------------------
		,(code		:= 17010
		,message 	:= '17010.  Start parameter for the compensation is invalid The section on which the compensation is to occur is not positive.')
		//318 -----------------------------------
		,(code		:= 17011
		,message 	:= '17011.  ?Target position under/overrun? (INTERNAL ERROR) The position (calculated from the modulo-target-position) where the axis should stand at end of oriented stop has been run over.')
		//319 -----------------------------------
		,(code		:= 17012
		,message 	:= '17012.  ?Target position will be under/overrun? (INTERNAL ERROR) The position (calculated from the modulo-target-position) where the axis should stand at end of oriented stop is too near and will be run over.')
		//320 -----------------------------------
		,(code		:= 17014
		,message 	:= '17014.  GROUPERR_GUIDERSTARTDATA')
		//321 -----------------------------------
		,(code		:= 17015
		,message 	:= '17015.  ?Dynamic parameters not permitted? (INTERNAL ERROR) The dynamic parameters resulting from internal calculation like acceleration, deceleration and jerk are not permitted.')
		//322 -----------------------------------
		,(code		:= 17017
		,message 	:= '17017.  GROUPERR_GUIDEROVERRUN')
		//323 -----------------------------------
		,(code		:= 17018
		,message 	:= '17018.  GROUPERR_GUIDERLOOKAHEAD')
		//324 -----------------------------------
		,(code		:= 17019
		,message 	:= '17019.  GROUPERR_GUIDERLOOKAHEADEND')
		//325 -----------------------------------
		,(code		:= 17020
		,message 	:= '17020.  GROUPERR_GUIDERLOOKAHEADREQU')
		//326 -----------------------------------
		,(code		:= 17021
		,message 	:= '17021.  GROUPERR_GUIDERMODE')
		//327 -----------------------------------
		,(code		:= 17022
		,message 	:= '17022.  ?A requested motion command could not be realized (BISECTION)? A requested motion command could not be realized using the requested parameters. The command has been executed best possible and this message is therefore to be understood just as a warning.')
		//328 -----------------------------------
		,(code		:= 17023
		,message 	:= '17023.  ?The new target position either has been overrun or will be overrun? The new target position either has been overrun or will be overrun, since until there it is impossible to stop. A internal stop command is commended.')
		//329 -----------------------------------
		,(code		:= 17024
		,message 	:= '17024.  Group not ready / group not ready for new task (INTERNAL ERROR / INFORMATION) The group is being given a new task while it is still in the process of executing an existing task. This request is not allowed because it would interrupt the execution of the previous task. The new task could, for instance, be a positioning command, or the set actual position function. Precisely the converse relationships apply for the set new end position function. In that case, the group/axis must still be actively moving in order to be able to cause a change in the end position.')
		//330 -----------------------------------
		,(code		:= 17025
		,message 	:= '17025.  The parameters of the oriented stop (O-Stop) are not admitted. The modulo-target position should not be smaller than zero and not larger or equal than the encoder mod-period ( e.g. in the interval [0.0,360.0) ).')
		//331 -----------------------------------
		,(code		:= 17026
		,message 	:= '17026.  The modulo target position of the modulo-start is invalid The modulo target position is outside of the valid parameter range. So the position value should not be smaller than zero and not greater or equal than the encoder modulo-period (e. g. in the interval [0.0,360.0) for the modulo starttype SHORTEST_WAY (261) ).')
		//332 -----------------------------------
		,(code		:= 17027
		,message 	:= '17027.  The online change activation mode is invalid. The activation can be used with online scaling or with online modification of motion function. The used activation is invalid in this context. Either the mode is not defined or yet not implemented or however it cannot in this constellation be put into action (e.g. when linear tables are used with an unexpected cyclic activation mode NEXTCYCLE or NEXTCYCLEONCE).')
		//333 -----------------------------------
		,(code		:= 17028
		,message 	:= '17028.  The parameterized jerk rate is not permitted. The jerk rate is smaller than the minimum jerk rate. The minimum value for jerk rate is 1.0 (e.g. mm/s^3).')
		//334 -----------------------------------
		,(code		:= 17029
		,message 	:= '17029.  The parameterized acceleration or deceleration is not permitted. The parameterized acceleration or deceleration is lower than the permitted minimum acceleration. The value for minimum acceleration is calculated from minimum jerk rate and NC cycle time (minimum jerk rate multiplied with NC cycle time). The unit for example is mm/s^2.')
		//335 -----------------------------------
		,(code		:= 17030
		,message 	:= '17030.  The parameterized velocity is not permitted. The parameterized target velocity is lower than the minimum velocity (but the value zero is permitted). The value for minimum velocity is calculated from the minimum jerk rate and the NC cycle time (minimum jerk rate multiplied with the square of the NC cycle time. The unit for example is mm/s.')
		//336 -----------------------------------
		,(code		:= 17031
		,message 	:= '17031.  A activation cannot be executed due to a pending activation A activation e.g. CamIn, CamScaling or WriteMotionFunction cannot be executed due to a pending activation (e.g. CamIn, CamScaling, WriteMotionFunction). Onle activation can be enabled.')
		//337 -----------------------------------
		,(code		:= 17032
		,message 	:= '17032.  ?Illegal combination of different cycle times within an axis group? A logical axis group includes elements (axes) with different cycle times for a common setpoint generator and I/O-execution, resp. This situation can occur with Master/Slave-coupling or configuring 3D- and FIFO-groups (including path, auxiliary, and slave axes).')
		//338 -----------------------------------
		,(code		:= 17033
		,message 	:= '17033.  Illegal motion reversal Due to the actual dynamical state a motion reversal will happen. To avoid this motion reversal the axis command is not performed and the previous system state restored.')
		//339 -----------------------------------
		,(code		:= 17034
		,message 	:= '17034.  ?Illegal moment for an axis command because there is an old axis command with activation position still active? The moment for the command is illegal because there is still an old command with activation position active (e.g. go to new velocity at threshold position or reach new velocity at threshold position).')
		//340 -----------------------------------
		,(code		:= 17035
		,message 	:= '17035.  Error in the stop-calculation routine (INTERNAL ERROR) Due to an internal error in the stop-calculation routine the current commando cannot be performed. The previous system state is restored.')
		//341 -----------------------------------
		,(code		:= 17036
		,message 	:= '17036.  A command with activation position cannot fully be performed because the remaining path is too short')
		//342 -----------------------------------
		,(code		:= 17037
		,message 	:= '17037.  Illegal decoupletype when decoupling a slave axis The decouple and restart command contains an invalid decouple type.')
		//343 -----------------------------------
		,(code		:= 17038
		,message 	:= '17038.  Illegal target velocity when decoupling a slave axis The decouple and restart command contains an illegal target velocity [1 < V <Vmax].')
		//344 -----------------------------------
		,(code		:= 17039
		,message 	:= '17039.  The command new dynamic parameter cannot be performed since this would require a new target velocity')
		//345 -----------------------------------
		,(code		:= 17040
		,message 	:= '17040.  ?A command with activation position cannot be performed becaus the axis is already in the brake phase?')
		//346 -----------------------------------
		,(code		:= 17041
		,message 	:= '17041.  ?Decouple routine of slave axis doesnt return a valid solution?')
		//347 -----------------------------------
		,(code		:= 17042
		,message 	:= '17042.  ?Command not be executed because the command buffer is full filled?')
		//348 -----------------------------------
		,(code		:= 17043
		,message 	:= '17043.  ?Command is rejected due to an internal error in the Look Ahead? (INTERNAL ERROR)')
		//349 -----------------------------------
		,(code		:= 17044
		,message 	:= '17044.  ?Command is rejected because the segment target velocity is not realized?')
		//350 -----------------------------------
		,(code		:= 17045
		,message 	:= '17045.  ?Successive commands have the same final position?')
		//351 -----------------------------------
		,(code		:= 17046
		,message 	:= '17046.  ?Logical positioning direction is inconsistent with the direction of the buffer command?')
		//352 -----------------------------------
		,(code		:= 17047
		,message 	:= '17047.  ?Command is rejected because the remaining positioning length is to small?')
		//353 -----------------------------------
		,(code		:= 17052
		,message 	:= '17052.  ?Reference cam is not found?  During the referencing process for an axis it is moved in the direction of the referencing cam. This reference cam, however, was not found as expected (=> leads to the abortion of the referencing procedure).')
		//354 -----------------------------------
		,(code		:= 17053
		,message 	:= '17053.  Reference cam became not free During the referencing process for an axis it is moved in the direction of the referencing cam, and is only stopped again when the cam signal is reached.  After the axis has also come to a physical standstill, the axis is subsequently started regularly from the cam again. In this case, the reference cam did not become free again as expected when driving down (=> leads to the abortion of the referencing procedure).')
		//355 -----------------------------------
		,(code		:= 17054
		,message 	:= '17054.  ?IO sync pulse was not found (only when using hardware latch)?. If the hardware latch is activated, a sync pulse (zero pulse) is expected to be found and a sync event triggered following the expiry of a certain time or a certain distance. If this is not the case, the reaction is an error and the abortion of the referencing procedure.')
		//356 -----------------------------------
		,(code		:= 17056
		,message 	:= '17056.  Group/axis consequential error Consequential error resulting from another causative error related to another axis within the group. Group/axis consequential errors can occur in relation to master/slave couplings or with multiple axis interpolating DXD groups. If, for instance, it is detected that the following error limit of a master axis has been exceeded, then this consequential error is assigned to all the other master axes and slave axes in this group.')
		//357 -----------------------------------
		,(code		:= 17057
		,message 	:= '17057.  Velocity reduction factor for C0/C1 transition is not allowed A C0 transition describes two geometries which, while they are themselves continuous, no not have either continuous first or second differentials. The velocity reduction factor C0 acts on such transitions.')
		//358 -----------------------------------
		,(code		:= 17058
		,message 	:= '17058.  Critical angle at segment transition not allowed')
		//359 -----------------------------------
		,(code		:= 17059
		,message 	:= '17059.  Radius of the tolerance sphere is in an invalid range')
		//360 -----------------------------------
		,(code		:= 17060
		,message 	:= '17060.  Not implemented.')
		//361 -----------------------------------
		,(code		:= 17061
		,message 	:= '17061.  Start type')
		//362 -----------------------------------
		,(code		:= 17062
		,message 	:= '17062.  Not implemented.')
		//363 -----------------------------------
		,(code		:= 17063
		,message 	:= '17063.  Blending with given parameters not possible')
		//364 -----------------------------------
		,(code		:= 17064
		,message 	:= '17064.  Not implemented.')
		//365 -----------------------------------
		,(code		:= 17065
		,message 	:= '17065.  Curve velocity reduction method not allowed (INTERNAL ERROR) The curve velocity reduction method does not exist.')
		//366 -----------------------------------
		,(code		:= 17066
		,message 	:= '17066.  Minimum velocity not allowed The minimum velocity that has been entered is less than 0.0.')
		//367 -----------------------------------
		,(code		:= 17067
		,message 	:= '17067.  Power function input not allowed (INTERNAL ERROR) The input parameters in the power_() function lead to an FPU exception.')
		//368 -----------------------------------
		,(code		:= 17068
		,message 	:= '17068.  Dynamic change parameter not allowed A parameter that controls alterations to the dynamics is invalid. parameters: 1. Absolute motion dynamics change: All parameters must be strictly positive. 2. Relative reduction c_f: 0.0 < c_f <= 1.0')
		//369 -----------------------------------
		,(code		:= 17069
		,message 	:= '17069.  Memory allocation error (INTERNAL ERROR)')
		//370 -----------------------------------
		,(code		:= 17070
		,message 	:= '17070.  The calculated end position differs from the end position in the nc instruction (internal error).')
		//371 -----------------------------------
		,(code		:= 17071
		,message 	:= '17071.  Calculate remaining chord length')
		//372 -----------------------------------
		,(code		:= 17072
		,message 	:= '17072.  Set value generator SVB active Starting the set value generator (SVB, SAF) has been refused, since the SVB task is already active.')
		//373 -----------------------------------
		,(code		:= 17073
		,message 	:= '17073.  SVB parameter not allowed (INTERNAL ERROR) A parameter related to the internal structure of the set value generator (SVB) results in logical errors and/or to an FPU exception. Affects these parameters: Minimum velocity (>0.0), TimeMode, ModeDyn, ModeGeo, StartType, DistanceToEnd, TBallRadius.')
		//374 -----------------------------------
		,(code		:= 17074
		,message 	:= '17074.  Velocity reduction factor not allowed A parameter that controls reduction of the velocity at segment transitions is invalid. Parameters: 1. Transitions with continuous first differential: VeloVertexFactorC1 2. Transitions without continuous differentials: VeloVertexFactorC0 CriticalVertexAngleLow, CriticalVertexAngleHigh.')
		//375 -----------------------------------
		,(code		:= 17075
		,message 	:= '17075.  Helix is a circle The helix has degenerated to a circle, and should be entered as such.')
		//376 -----------------------------------
		,(code		:= 17076
		,message 	:= '17076.  Helix is a straight line The helix has degenerated to a straight line, and should be entered as such.')
		//377 -----------------------------------
		,(code		:= 17077
		,message 	:= '17077.  Guider parameter not allowed One of the guiders parameters leads to logical errors and/or to an FPU exception.')
		//378 -----------------------------------
		,(code		:= 17078
		,message 	:= '17078.  Invalid segment address (INTERNAL ERROR) The geometry segment does not have a valid geometry structure address or does not have a valid dynamic structure address.')
		//379 -----------------------------------
		,(code		:= 17079
		,message 	:= '17079.  Unparametrised generator (INTERNAL ERROR) The SVB generator is not yet parameterised and is therefore unable to operate.')
		//380 -----------------------------------
		,(code		:= 17080
		,message 	:= '17080.  Unparametrised table (INTERNAL ERROR) The table has no information concerning the address of the corresponding dynamic generator.')
		//381 -----------------------------------
		,(code		:= 17082
		,message 	:= '17082.  The calculation of the arc length of the smoothed path failed (internal error).')
		//382 -----------------------------------
		,(code		:= 17083
		,message 	:= '17083.  The radius of the tolerance ball is too small (smaller than 0.1 mm).')
		//383 -----------------------------------
		,(code		:= 17084
		,message 	:= '17084.  Error while calculating DXD-Software-Limitswitches (internal error))')
		//384 -----------------------------------
		,(code		:= 17085
		,message 	:= '17085.  NC-Block violates software limit switches of the group At least one path axis with active software limit monitoring has violated the limit switches Therefore the geometric entry is denied with an error.')
		//385 -----------------------------------
		,(code		:= 17086
		,message 	:= '17086.  GROUPERR_DXD_SOFTENDCHECK')
		//386 -----------------------------------
		,(code		:= 17087
		,message 	:= '17087.  GROUPERR_DXD_RTTG_VELOREFERENCE')
		//387 -----------------------------------
		,(code		:= 17088
		,message 	:= '17088.  Interpolating group contains axes of an incorrect axis type An interpolating 3D group may only contain continuously guided axes of axis type 1 (SERVO).')
		//388 -----------------------------------
		,(code		:= 17089
		,message 	:= '17089.  Scalar product can not be calculated The length of one of the given vectors is 0.0.')
		//389 -----------------------------------
		,(code		:= 17090
		,message 	:= '17090.  Inverse cosine can not be calculated The length of one of the given vectors is 0.0.')
		//390 -----------------------------------
		,(code		:= 17091
		,message 	:= '17091.  Invalid table entry type The given table entry type is unknown.')
		//391 -----------------------------------
		,(code		:= 17092
		,message 	:= '17092.  Invalid DIN66025 information type (INTERNAL ERROR) The given DIN66025 information type is unknown. Known types: G0, G1, G2, G3, G17, G18, G19.')
		//392 -----------------------------------
		,(code		:= 17093
		,message 	:= '17093.  Invalid dimension (INTERNAL ERROR) The CNC dimension is unknown. Known dimensions: 1, 2, 3. Or: The CNC dimension is invalid for the given geometrical object. For a circle the dimension must be 2 or 3, while for a helix it must be 3.')
		//393 -----------------------------------
		,(code		:= 17094
		,message 	:= '17094.  Geometrical object is not a straight line The given object, interpreted as a straight line, has a length of 0.0.')
		//394 -----------------------------------
		,(code		:= 17095
		,message 	:= '17095.  Geometrical object is not a circle Interpreted as a circular arc, the given object has a length of 0.0, or an angle of 0.0 or a radius of 0.0.')
		//395 -----------------------------------
		,(code		:= 17096
		,message 	:= '17096.  Geometrical object is not a helix Interpreted as a circular arc, the given object has a length of 0.0, or an angle of 0.0, or a radius of 0.0. or a height of 0.0.')
		//396 -----------------------------------
		,(code		:= 17097
		,message 	:= '17097.  Set velocity less than or equal to 0.0 is invalid A value less than or equal to 0.0 for the set velocity (CNC) is not allowed, since the set velocity is positive by definition, and a set velocity of 0.0 cannot generate any motion.')
		//397 -----------------------------------
		,(code		:= 17098
		,message 	:= '17098.  Address for look-ahead invalid (INTERNAL ERROR) The address supplied for the look-ahead is invalid.')
		//398 -----------------------------------
		,(code		:= 17099
		,message 	:= '17099.  Set value generator SAF active Starting the set value generator (SAF) has been refused, since the SAF task is already active.')
		//399 -----------------------------------
		,(code		:= 17100
		,message 	:= '17100.  CNC set value generation not active Stop or change of override refused, because the set value generation is not active.')
		//400 -----------------------------------
		,(code		:= 17101
		,message 	:= '17101.  CNC set value generation in the stop phase Stop or change of override refused, because the set value generation is in the stop phase.')
		//401 -----------------------------------
		,(code		:= 17102
		,message 	:= '17102.  Override not allowed An override of less than 0.0% or more than 100.0% is invalid.')
		//402 -----------------------------------
		,(code		:= 17103
		,message 	:= '17103.  Invalid table address (INTERNAL ERROR) The table address given for the initialisation of the set value generator is invalid, or no valid logger connection (report file) is present.')
		//403 -----------------------------------
		,(code		:= 17104
		,message 	:= '17104.  Invalid table entry type The given table entry type is unknown.')
		//404 -----------------------------------
		,(code		:= 17105
		,message 	:= '17105.  Memory allocation failed Memory allocation for the table has failed.')
		//405 -----------------------------------
		,(code		:= 17106
		,message 	:= '17106.  Memory allocation failed Memory allocation for the filter has failed.')
		//406 -----------------------------------
		,(code		:= 17107
		,message 	:= '17107.  Invalid parameter Filter parameter is not allowed.')
		//407 -----------------------------------
		,(code		:= 17108
		,message 	:= '17108.  Delete Distance To Go failed Delete Distance to go (only interpolation) failed. This error occured, if e.g. the command DelDTG was not programmed in the actual movement of the nc program.')
		//408 -----------------------------------
		,(code		:= 17109
		,message 	:= '17109.  The setpoint generator of the fying saw generates incompatible values (internal error)')
		//409 -----------------------------------
		,(code		:= 17110
		,message 	:= '17110.  Axis will be stopped since otherwise it will overrun its target position (old PTP setpoint generator) If, for example, in case of a slave to master transformation for the new master a target position is commanded that will be overrun because of the actual dynamics the axis will be stopped internally to guarantee that the target position will not be overrun.')
		//410 -----------------------------------
		,(code		:= 17111
		,message 	:= '17111.  Internal error in the transformation from slave to master.')
		//411 -----------------------------------
		,(code		:= 17112
		,message 	:= '17112.  Wrong direction in the transformation of slave to master.')
		//412 -----------------------------------
		,(code		:= 17114
		,message 	:= '17114.  Parameter of Motion Function (MF) table incorrect The parameter of the Motion Function (MF) are incorrect. This may refer to the first time created data set or to online changed data.')
		//413 -----------------------------------
		,(code		:= 17115
		,message 	:= '17115.  Parameter of Motion Function (MF) table incorrect The parameter of the Motion Function (MF) are invalid. This may refer to the first time created data set or to online changed data. The error cause can be, that an active MF point (no IGNORE point) points at a passive MF point (IGNORE point).')
		//414 -----------------------------------
		,(code		:= 17116
		,message 	:= '17116.  Internal error by using Motion Function (MF) An internal error occurs by using the Function (MF). This error can not be solved by the user. Plaese ask the TwinCAT Support.')
		//415 -----------------------------------
		,(code		:= 17117
		,message 	:= '17117.  Axis coupling with synchronization generator declined because of incorrect axis dynamic values The axis coupling with the synchronization generator has been declined, because one of the slave dynamic parameter (machine data) is incorrect (e.g. the maximum velocity, the acceleration, the deceleration or the jerk is smaller or equal to zero, or the expected synchronous velocity of the slave axis is higher as the maximum allowed slave velocity.')
		//416 -----------------------------------
		,(code		:= 17118
		,message 	:= '17118.  Coupling conditions of synchronization generator incorrect')
		//417 -----------------------------------
		,(code		:= 17119
		,message 	:= '17119.  Moving profile of synchronization generator declines dynamic limit of slave axis or required characterstic of profile One of the parameterized checks has recognized an overstepping of the dynamic limits (max. velocity, max. acceleration, max. deceleration or max. jerk) of the slave axis, or an profile characteristic (e.g. overshoot or undershoot in the position or velocity) is incorrect. See also further messages in the windows event log and in the message window of the System Manager.')
		//418 -----------------------------------
		,(code		:= 17120
		,message 	:= '17120.  Invalid parameter The encoder generator parameter is not allowed.')
		//419 -----------------------------------
		,(code		:= 17121
		,message 	:= '17121.  Invalid parameter The external (Fifo) generator parameter is not allowed.')
		//420 -----------------------------------
		,(code		:= 17122
		,message 	:= '17122.  External generator is active The external generator cannot be started, as it is already active.')
		//421 -----------------------------------
		,(code		:= 17123
		,message 	:= '17123.  External generator is not active The external generator cannot be stopped, as it is not active.')
		//422 -----------------------------------
		,(code		:= 17124
		,message 	:= '17124.  NC-Block with auxiliary axis violates software limit switches of the group At least one auxiliary axis with active software limit monitoring has violated the limit switches Therefore the geometric entry is denied with an error.')
		//423 -----------------------------------
		,(code		:= 17125
		,message 	:= '17125.  NC-Block type Bezier spline curve contains a cusp (singularity) The Bezier spline curve contain a cusp, i.e. at a certain interior point both the curvature and the modulus of the velocity tend to 0 such that the radius of curvature is infinite.')
		//424 -----------------------------------
		,(code		:= 17127
		,message 	:= '17127.  ?Value for dead time compensation not allowed? The value for the dead time compensation in seconds for a slave coupling to an encoder axis (virtual axis) is not allowed.')
		//425 -----------------------------------
		,(code		:= 17128
		,message 	:= '17128.  GROUPERR_RANGE_NOMOTIONWINDOW')
		//426 -----------------------------------
		,(code		:= 17129
		,message 	:= '17129.  GROUPERR_RANGE_NOMOTIONFILTERTIME')
		//427 -----------------------------------
		,(code		:= 17130
		,message 	:= '17130.  GROUPERR_RANGE_TIMEUNITFIFO')
		//428 -----------------------------------
		,(code		:= 17131
		,message 	:= '17131.  GROUPERR_RANGE_OVERRIDETYPE')
		//429 -----------------------------------
		,(code		:= 17132
		,message 	:= '17132.  GROUPERR_RANGE_OVERRIDECHANGETIME')
		//430 -----------------------------------
		,(code		:= 17133
		,message 	:= '17133.  GROUPERR_FIFO_INVALIDDIMENSION')
		//431 -----------------------------------
		,(code		:= 17134
		,message 	:= '17134.  GROUPERR_ADDR_FIFOTABLE')
		//432 -----------------------------------
		,(code		:= 17135
		,message 	:= '17135.  Axis is locked for motion commands because a stop command is still activeThe axis/group is locked for motion commands because a stop command is still active. The axis can be released by calling MC_Stop with Execute=FALSE or by using MC_Reset (TcMC2.Lib).')
		//433 -----------------------------------
		,(code		:= 17136
		,message 	:= '17136.  Invalid number of auxiliary axes The local number of auxiliary axes does not tally with the global number of auxiliary axes.')
		//434 -----------------------------------
		,(code		:= 17137
		,message 	:= '17137.  Invalid reduction parameter for auxiliary axes The velocity reduction parameters for the auxiliary axes are inconsistent.')
		//435 -----------------------------------
		,(code		:= 17138
		,message 	:= '17138.  Invalid dynamic parameter for auxiliary axes The dynamic parameters for the auxiliary axes are inconsistent.')
		//436 -----------------------------------
		,(code		:= 17139
		,message 	:= '17139.  Invalid coupling parameter for auxiliary axes The coupling parameters for the auxiliary axes are inconsistent.')
		//437 -----------------------------------
		,(code		:= 17140
		,message 	:= '17140.  Invalid auxiliary axis entry The auxiliary axis entry is empty (no axis motion).')
		//438 -----------------------------------
		,(code		:= 17142
		,message 	:= '17142.  Invalid parameter The limit for velocity reduction of the auxiliary axes is invalid. It has to be in the interval 0..1.0')
		//439 -----------------------------------
		,(code		:= 17151
		,message 	:= '17151.  GROUPERR_HYMMEN_WATCHDOG')
		//440 -----------------------------------
		,(code		:= 17152
		,message 	:= '17152.  Axis ID not allowed The value for the axis ID is not allowed, e.g. because it has already been assigned, is less than or equal to zero, is greater than 255, or does not exist in the current configuration.')
		//441 -----------------------------------
		,(code		:= 17153
		,message 	:= '17153.  Axis type not allowed The value for the axis type is unacceptable because it is not defined. Type 1: Servo Type 2: High/low speed Type 3: Stepper motor')
		//442 -----------------------------------
		,(code		:= 17158
		,message 	:= '17158.  Slow manual velocity not allowed The value for the slow manual velocity is not allowed.')
		//443 -----------------------------------
		,(code		:= 17159
		,message 	:= '17159.  Fast manual velocity not allowed The value for the fast manual velocity is not allowed.')
		//444 -----------------------------------
		,(code		:= 17160
		,message 	:= '17160.  High speed not allowed The value for the high speed is not allowed.')
		//445 -----------------------------------
		,(code		:= 17161
		,message 	:= '17161.  Acceleration not allowed The value for the axis acceleration is not allowed.')
		//446 -----------------------------------
		,(code		:= 17162
		,message 	:= '17162.  Deceleration not allowed The value for the axis deceleration is not allowed.')
		//447 -----------------------------------
		,(code		:= 17163
		,message 	:= '17163.  Jerk not allowed The value for the axis jerk is not allowed.')
		//448 -----------------------------------
		,(code		:= 17164
		,message 	:= '17164.  Delay time between position and velocity is not allowed The value for the delay time between position and velocity (idle time compensation) is not allowed.')
		//449 -----------------------------------
		,(code		:= 17165
		,message 	:= '17165.  ?Override-Type not allowed? The value for the velocity override type is not allowed. Type 1: With respect to the internal reduced velocity (default value) Type 2: With respect to the original external start velocity')
		//450 -----------------------------------
		,(code		:= 17166
		,message 	:= '17166.  NCI: Velo-Jump-Factor not allowed')
		//451 -----------------------------------
		,(code		:= 17167
		,message 	:= '17167.  NCI: Radius of tolerance sphere for the auxiliary axes is invalid')
		//452 -----------------------------------
		,(code		:= 17168
		,message 	:= '17168.  NCI: Value for maximum deviation for the auxiliary axes is invalid')
		//453 -----------------------------------
		,(code		:= 17170
		,message 	:= '17170.  Referencing velocity in direction of cam not allowed The value for the referencing velocity in the direction of the referencing cam is not allowed.')
		//454 -----------------------------------
		,(code		:= 17171
		,message 	:= '17171.  Referencing velocity in sync direction not allowed The value for the referencing velocity in the direction of the sync pulse (zero track) is not allowed.')
		//455 -----------------------------------
		,(code		:= 17172
		,message 	:= '17172.  Pulse width in positive direction not allowed The value for the pulse width in the positive direction is not allowed (pulsed operation). The use of the pulse width for positioning is chosen implicitly through the axis start type. Pulsed operation corresponds to positioning with a relative displacement that corresponds precisely to the pulse width.')
		//456 -----------------------------------
		,(code		:= 17173
		,message 	:= '17173.  Pulse width in negative direction not allowed The value for the pulse width in the negative direction is not allowed (pulsed operation). The use of the pulse width for positioning is chosen implicitly through the axis start type. Pulsed operation corresponds to positioning with a relative displacement that corresponds precisely to the pulse width.')
		//457 -----------------------------------
		,(code		:= 17174
		,message 	:= '17174.  Pulse time in positive direction not allowed The value for the pulse width in the positive direction is not allowed (pulsed operation).')
		//458 -----------------------------------
		,(code		:= 17175
		,message 	:= '17175.  Pulse time in negative direction not allowed The value for the pulse width in the negative direction is not allowed (pulsed operation).')
		//459 -----------------------------------
		,(code		:= 17176
		,message 	:= '17176.  Creep distance in positive direction not allowed The value for the creep distance in the positive direction is not allowed.')
		//460 -----------------------------------
		,(code		:= 17177
		,message 	:= '17177.  Creep distance in negative direction not allowed The value for the creep distance in the negative direction is not allowed.')
		//461 -----------------------------------
		,(code		:= 17178
		,message 	:= '17178.  Braking distance in positive direction not allowed The value for the braking distance in the positive direction is not allowed.')
		//462 -----------------------------------
		,(code		:= 17179
		,message 	:= '17179.  Braking distance in negative direction not allowed The value for the braking distance in the negative direction is not allowed.')
		//463 -----------------------------------
		,(code		:= 17180
		,message 	:= '17180.  Braking time in positive direction not allowed The value for the braking time in the positive direction is not allowed.')
		//464 -----------------------------------
		,(code		:= 17181
		,message 	:= '17181.  Braking time in negative direction not allowed The value for the braking time in the negative direction is not allowed.')
		//465 -----------------------------------
		,(code		:= 17182
		,message 	:= '17182.  Switching time from high to low speed not allowed The value for the time to switch from high to low speed is not allowed.')
		//466 -----------------------------------
		,(code		:= 17183
		,message 	:= '17183.  Creep distance for stop not allowed The value for the creep distance for an explicit stop is not allowed.')
		//467 -----------------------------------
		,(code		:= 17184
		,message 	:= '17184.  Motion monitoring not allowed The value for the activation of the motion monitoring is not allowed.')
		//468 -----------------------------------
		,(code		:= 17185
		,message 	:= '17185.  Position window monitoring not allowed The value for the activation of the position window monitoring is not allowed.')
		//469 -----------------------------------
		,(code		:= 17186
		,message 	:= '17186.  Target window monitoring not allowed The value for the activation of target window monitoring is not allowed.')
		//470 -----------------------------------
		,(code		:= 17187
		,message 	:= '17187.  Loop not allowed The value for the activation of loop movement is not allowed.')
		//471 -----------------------------------
		,(code		:= 17188
		,message 	:= '17188.  Motion monitoring time not allowed The value for the motion monitoring time is not allowed.')
		//472 -----------------------------------
		,(code		:= 17189
		,message 	:= '17189.  Target window range not allowed The value for the target window is not allowed.')
		//473 -----------------------------------
		,(code		:= 17190
		,message 	:= '17190.  Position window range not allowed The value for the position window is not allowed.')
		//474 -----------------------------------
		,(code		:= 17191
		,message 	:= '17191.  Position window monitoring time not allowed The value for the position window monitoring time is not allowed.')
		//475 -----------------------------------
		,(code		:= 17192
		,message 	:= '17192.  Loop movement not allowed The value for the loop movement is not allowed.')
		//476 -----------------------------------
		,(code		:= 17193
		,message 	:= '17193.  Axis cycle time not allowed The value for the axis cycle time is not allowed.')
		//477 -----------------------------------
		,(code		:= 17194
		,message 	:= '17194.  Stepper motor operating mode not allowed The value for the stepper motor operating mode is not allowed.')
		//478 -----------------------------------
		,(code		:= 17195
		,message 	:= '17195.  Displacement per stepper motor step not allowed The value for the displacement associated with one step of the stepper motor is not allowed (step scaling). Value range: [0.000001, 1000.0]                                     Unit: e.g. mm/STEP')
		//479 -----------------------------------
		,(code		:= 17196
		,message 	:= '17196.  Minimum speed for stepper motor set value profile not allowed The value for the minimum speed of the stepper motor speed profile is not allowed.')
		//480 -----------------------------------
		,(code		:= 17197
		,message 	:= '17197.  Stepper motor stages for one speed stage not allowed The value for the number of steps for each speed stage in the set value generation is not allowed.')
